// TIA Portal V21 export
// export: Created 2026-11-18T11:11:29.3256104Z, ExportSetting WithDefaults, DisplayName Totally Integrated Automation Portal, DisplayVersion V21, DisplayName STEP 7 Professional, DisplayVersion V21, DisplayName STEP 7 Safety, DisplayVersion V21, DisplayName Tech WebApplication, DisplayVersion V21, DisplayName WinCC Basic/Comfort/Advanced, DisplayVersion V21
Screen "Screen_Template"  800x480, Number=2
  ScreenLayer 
    Circle "Circle_1" at 39,39 size 48x48
      RangeAppearanceAnimation "RangeAppearanceAnimation"
        tag PLC_Sys_Status
        0..0: back #dedbde, fore #181c31
        1..1: back #00ff00, fore #181c31
        2..2: back #ff0000, fore #181c31, flashing
    TextField "Text field_1" at 177,40 size 43x23  Text="Text"
      VisibilityAnimation "VisibilityAnimation"  RangeEnd=1
        tag PLC_Alm_Missing_Prod
    IOField "I/O field_1" at 267,46 size 96x32  DataFormat=Decimal, FormatPattern=9999999, Mode=Output
      ProcessValue := PLC_Cognex_Sensor_Count
    Button "Button_1" at 425,46 size 150x32  Mode=Text, TextOff="HMI_Btn_Start;", TextOn="Text"
      on Press: SetBit(Tag := HMI_Btn_Start)
      on Release: ResetBit(Tag := HMI_Btn_Start)
    Button "Button_2" at 426,119 size 186x32  Mode=Text, TextOff="HMI_Sw_Mode_Auto.", TextOn="Text"
      on Click: InvertBit(Tag := HMI_Sw_Mode_Auto)
